Fanuc KAREL source: kt00891.KL

-- PROVISIONAL review KL for V940-1; original PC SHA256 683b6cc714d7d8809d105a70be03aa367a1432563352916909cbb39c62e45bc1
-- Incomplete behavior may be omitted. Consult companion uncertainty JSON. Do not deploy.
PROGRAM KT00891
%NOLOCKGROUP
-- UNRESOLVED_DECL P1 type=000199
-- UNRESOLVED_DECL P2 type=000199
-- UNRESOLVED_DECL OUT type=000101
BEGIN
  -- V9_ZERO_TABLE_METADATA_HINT layout=0001; no indexed target words; source/name/runtime held
  -- UNRESOLVED_PC offsets 5-35; opcodes 27,27,49,7E,AD,76,7E,4A
  -- UNRESOLVED_PC offsets 40-44; opcodes 7F
END KT00891
